Fanuc TP program (LS listing): DropEa.LS

/PROG  DropEa
/ATTR
OWNER		= MNEDITOR;
COMMENT		= "RoboDK sequence";
PROG_SIZE	= 0;
CREATE		= DATE 31-12-14  TIME 12:00:00;
MODIFIED	= DATE 31-12-14  TIME 12:00:00;
FILE_NAME	= DropEa;
VERSION		= 0;
LINE_COUNT	= 23;
MEMORY_SIZE	= 0;
PROTECT		= READ_WRITE;
TCD:  STACK_SIZE	= 0,
      TASK_PRIORITY	= 50,
      TIME_SLICE	= 0,
      BUSY_LAMP_OFF	= 0,
      ABORT_REQUEST	= 0,
      PAUSE_REQUEST	= 0;
DEFAULT_GROUP	= 1,*,*,*,*;
CONTROL_CODE	= 00000000 00000000;
/MN
   1:  ! Program generated by VerticalBot Studio for Fanuc LR Mate 200 ;
   2:  ! iD/7L on 25/10/2026 12:00:00 ;
   3:  ! Using nominal kinematics. ;
   4:  PR[9,1]=160.000 ;
   5:  PR[9,2]=-540.000 ;
   6:  PR[9,3]=300.000 ;
   7:  PR[9,4]=0.000 ;
   8:  PR[9,5]=0.000 ;
   9:  PR[9,6]=-180.000 ;
  10:  UFRAME[9]=PR[9] ;
  11:  UFRAME_NUM=9 ;
  12:  PR[9,1]=0.000 ;
  13:  PR[9,2]=0.000 ;
  14:  PR[9,3]=70.000 ;
  15:  PR[9,4]=0.000 ;
  16:  PR[9,5]=0.000 ;
  17:  PR[9,6]=0.000 ;
  18:  UTOOL[9]=PR[9] ;
  19:  UTOOL_NUM=9 ;
  20:J P[1] 20% FINE ;
  21:L P[2] 200mm/sec FINE ;
  22:  CALL Drop ;
  23:J P[3] 20% FINE ;
/POS
P[1]{
   GP1:
    UF : 9, UT : 9,
	J1=    -40.156 deg,	J2=    -35.956 deg,	J3=    -12.422 deg,
	J4=    100.287 deg,	J5=    -50.967 deg,	J6=    -16.077 deg
};
P[2]{
   GP1:
    UF : 9, UT : 9,        CONFIG : 'F U T, 0, 0, 0',
	X =     0.000  mm,	Y =    75.000  mm,	Z =     0.000  mm,
	W =    90.000 deg,	P =     0.000 deg,	R =  -180.000 deg
};
P[3]{
   GP1:
    UF : 9, UT : 9,
	J1=    -40.156 deg,	J2=    -35.956 deg,	J3=    -12.422 deg,
	J4=    100.287 deg,	J5=    -50.967 deg,	J6=    -16.077 deg
};
/END
